(* IEC 61131-3 sources: teller/JD_Teller_LC2_V11/Network/Teller, 1 file *)

(* ---- ONE_Teller_Table.st ---- *)
#define OBJECTS_CONFIG

FUNCTION GLOBAL TAB ONE_Teller
-1$UINT, 0$UINT,
0$UINT, 0$UINT,

13$UDINT,
TO_UDINT(3073024365), "Encoder_Inmeten", 0$UINT, 0$UINT, 1$UINT,
TO_UDINT(1689253198), "FileBase", 1$UINT, 0$UINT, 2$UINT,
TO_UDINT(2225119864), "MerkerEx", 1$UINT, 18$UINT, 2$UINT,
TO_UDINT(1903583397), "Ram", 1$UINT, 3$UINT, 16$UINT,
TO_UDINT(933570811), "RAMex", 1$UINT, 16$UINT, 1$UINT,
TO_UDINT(582296389), "SerSend", 1$UINT, 0$UINT, 1$UINT,
TO_UDINT(1018833242), "SIMPULSJE_Teller", 1$UINT, 0$UINT, 1$UINT,
TO_UDINT(1850111279), "String", 1$UINT, 10$UINT, 2$UINT,
TO_UDINT(2898603620), "StringInternal", 1$UINT, 70$UINT, 0$UINT,
TO_UDINT(2685101138), "TanabeCounterSerial", 1$UINT, 0$UINT, 1$UINT,
TO_UDINT(4092741209), "TellerClass_Teller", 1$UINT, 3$UINT, 1$UINT,
TO_UDINT(3232495061), "VirtualBaseInit", 1$UINT, 3$UINT, 0$UINT,
TO_UDINT(589051502), "VisuTeller_Teller", 1$UINT, 0$UINT, 5$UINT,

_NO_ATTR, TO_UDINT(2959661299), "ENCODER_INMETEN1",

_NO_ATTR, TO_UDINT(316419285), "FILEBASE1",
_NO_ATTR, TO_UDINT(2346024303), "FILEBASE2",

1$UINT, TO_UDINT(3025948), "STRING1\MERKEREX0",
1$UINT, TO_UDINT(1480758749), "STRING3\MERKEREX0",

1$UINT, TO_UDINT(4072236793), "SERSEND1\RSELECTOR",
1$UINT, TO_UDINT(3232725082), "TELLERCLASS1\RI2SENCNT",
1$UINT, TO_UDINT(3756668069), "TELLERCLASS1\RIBOXLENGTHCNT",
1$UINT, TO_UDINT(3865050826), "TELLERCLASS1\RIBOXLENGTHJAML",
1$UINT, TO_UDINT(475055017), "TELLERCLASS1\RIBOXLENGTHJAMR",
1$UINT, TO_UDINT(1711364282), "TELLERCLASS1\RIBOXLENGTHJAMSTR",
1$UINT, TO_UDINT(1431716753), "TELLERCLASS1\RIENCDIV",
1$UINT, TO_UDINT(1100143673), "TELLERCLASS1\RIENCMUL",
1$UINT, TO_UDINT(3615109569), "TELLERCLASS1\RISENSORCNT",
1$UINT, TO_UDINT(1331113651), "TELLERCLASS1\RITOTALPRODUCTION",
1$UINT, TO_UDINT(632896864), "TELLERCLASS1\RMINSPOT",
1$UINT, TO_UDINT(1272264235), "TELLERCLASS1\ROCOUNTER",
1$UINT, TO_UDINT(1448788453), "TELLERCLASS1\RSANALOGSPEEDENABLE",
1$UINT, TO_UDINT(3322901645), "TELLERCLASS1\RSEXTRABOX",
1$UINT, TO_UDINT(2626903235), "TELLERCLASS1\RSFACTORANALOGSPEEDIN",
1$UINT, TO_UDINT(2919943508), "TELLERCLASS1\RSMAXSPEED",

_NO_ATTR, TO_UDINT(1200226343), "RAMEX3",

_NO_ATTR, TO_UDINT(2236149643), "SERSEND1",

_NO_ATTR, TO_UDINT(3969721823), "SIMPULSJE5",

_NO_ATTR, TO_UDINT(677614747), "STRING1",
_NO_ATTR, TO_UDINT(3329095095), "STRING3",

_NO_ATTR, TO_UDINT(3886509187), "READ_SERIAL1",

_NO_ATTR, TO_UDINT(326458637), "TELLERCLASS1",

_NO_ATTR, TO_UDINT(2767617665), "VISUTELLER1",
_NO_ATTR, TO_UDINT(1040133947), "VISUTELLER2",
_NO_ATTR, TO_UDINT(1257775021), "VISUTELLER3",
_NO_ATTR, TO_UDINT(3567028750), "VISUTELLER4",
_NO_ATTR, TO_UDINT(2744892056), "VISUTELLER5",

//Internal connections
0$UDINT,
18$UDINT,
TO_UDINT(22), "rSelector", TO_UDINT(5),
TO_UDINT(24), "MerkerEx0", TO_UDINT(3),
TO_UDINT(25), "MerkerEx0", TO_UDINT(4),
TO_UDINT(27), "RMinSpot", TO_UDINT(15),
TO_UDINT(27), "rSextraBox", TO_UDINT(18),
TO_UDINT(27), "riEncMul", TO_UDINT(12),
TO_UDINT(27), "riEncDiv", TO_UDINT(11),
TO_UDINT(27), "riSensorCNT", TO_UDINT(13),
TO_UDINT(27), "riBoxlengthCNT", TO_UDINT(7),
TO_UDINT(27), "riTotalProduction", TO_UDINT(14),
TO_UDINT(27), "riBoxlengthJAML", TO_UDINT(8),
TO_UDINT(27), "riBoxlengthJAMR", TO_UDINT(9),
TO_UDINT(27), "riBoxlengthJamSTR", TO_UDINT(10),
TO_UDINT(27), "roCounter", TO_UDINT(16),
TO_UDINT(27), "ri2SenCNT", TO_UDINT(6),
TO_UDINT(27), "rsMaxSpeed", TO_UDINT(20),
TO_UDINT(27), "rsFactorAnalogSpeedIn", TO_UDINT(19),
TO_UDINT(27), "rsAnalogSpeedEnable", TO_UDINT(17),
0$UDINT,
27$UDINT,
TO_UDINT(22), "fb", TO_UDINT(1), "Server0",
TO_UDINT(22), "strSend", TO_UDINT(25), "Data",
TO_UDINT(24), "DataBuffer", TO_UDINT(3), "m_udLength",
TO_UDINT(25), "DataBuffer", TO_UDINT(4), "m_udLength",
TO_UDINT(26), "GetInfo", TO_UDINT(27), "ClassSvr",
TO_UDINT(26), "String", TO_UDINT(24), "Data",
TO_UDINT(26), "FileBase", TO_UDINT(2), "Server0",
TO_UDINT(26), "cPlannedProduction", TO_UDINT(27), "iTotalProduction",
TO_UDINT(26), "cBoxLength", TO_UDINT(27), "iBoxlengthCNT",
TO_UDINT(26), "cBattingStart", TO_UDINT(30), "iStart",
TO_UDINT(26), "cBattingDistance", TO_UDINT(30), "iLengte",
TO_UDINT(26), "cBatch1", TO_UDINT(30), "iPakket1SET",
TO_UDINT(26), "cBatch2", TO_UDINT(30), "iPakket2SET",
TO_UDINT(26), "cStartingDistanceToConveyorRun", TO_UDINT(29), "iLengte",
TO_UDINT(26), "cCountedBoxes", TO_UDINT(27), "oCounter",
TO_UDINT(27), "RamEx", TO_UDINT(21), "m_udLength",
TO_UDINT(27), "iSimPuls", TO_UDINT(23), "Uitgang",
TO_UDINT(27), "coTotalproduction", TO_UDINT(22), "iTotalproduction",
TO_UDINT(27), "coCounter", TO_UDINT(22), "iCounter",
TO_UDINT(27), "coRemainingproduction", TO_UDINT(22), "iRemaningproduction",
TO_UDINT(27), "coCounterPerMin", TO_UDINT(22), "iCounterPerMin",
TO_UDINT(27), "coSpeed", TO_UDINT(22), "iSpeed",
TO_UDINT(28), "cData", TO_UDINT(27), "sData",
TO_UDINT(29), "cData", TO_UDINT(27), "sData",
TO_UDINT(30), "cData", TO_UDINT(27), "sData",
TO_UDINT(31), "cData", TO_UDINT(27), "sData",
TO_UDINT(32), "cData", TO_UDINT(27), "sData",

//Initialization values
0$UDINT,
19$UDINT,
TO_UDINT(0), "cEncoder", TO_UDINT(0),//|Teller.Encoder_Inmeten1.cEncoder;
TO_UDINT(3), "ThreadSafe", TO_UDINT(0),//|Teller.String1\MerkerEx0.ThreadSafe;
TO_UDINT(4), "ThreadSafe", TO_UDINT(0),//|Teller.String3\MerkerEx0.ThreadSafe;
TO_UDINT(21), "ThreadSafe", TO_UDINT(0),//|Teller.RAMex3.ThreadSafe;
TO_UDINT(24), "SingleRealloc", TO_UDINT(1),//|Teller.String1.SingleRealloc;
TO_UDINT(26), "GetInfo", TO_UDINT(0),//|Teller.Read_serial1.GetInfo;
TO_UDINT(27), "iSensorSTR", TO_UDINT(0),//|Teller.TellerClass1.iSensorSTR;
TO_UDINT(27), "oJam", TO_UDINT(0),//|Teller.TellerClass1.oJam;
TO_UDINT(27), "cExtBoxCount", TO_UDINT(0),//|Teller.TellerClass1.cExtBoxCount;
TO_UDINT(28), "cHeadNr", TO_UDINT(1),//|Teller.VisuTeller1.cHeadNr;
TO_UDINT(28), "cType", TO_UDINT(4),//|Teller.VisuTeller1.cType;
TO_UDINT(29), "cHeadNr", TO_UDINT(2),//|Teller.VisuTeller2.cHeadNr;
TO_UDINT(29), "cType", TO_UDINT(3),//|Teller.VisuTeller2.cType;
TO_UDINT(30), "cHeadNr", TO_UDINT(3),//|Teller.VisuTeller3.cHeadNr;
TO_UDINT(30), "cType", TO_UDINT(1),//|Teller.VisuTeller3.cType;
TO_UDINT(31), "cHeadNr", TO_UDINT(4),//|Teller.VisuTeller4.cHeadNr;
TO_UDINT(31), "cType", TO_UDINT(5),//|Teller.VisuTeller4.cType;
TO_UDINT(32), "cHeadNr", TO_UDINT(5),//|Teller.VisuTeller5.cHeadNr;
TO_UDINT(32), "cType", TO_UDINT(2),//|Teller.VisuTeller5.cType;

//Symbolic initialization values
0$UDINT,
0$UDINT,

//Initialization of string values
0$UDINT,
0$UDINT,

//Configuration of tasks (RealTime, Cyclic, Background)
0$UDINT,
1$UDINT,
TO_UDINT(27), (1)$UDINT, 4194305$DINT, 	//TELLERCLASS1

0$UDINT,
3$UDINT,
TO_UDINT(26), (1)$UDINT, 4194303$DINT, 	//READ_SERIAL1
TO_UDINT(23), (10)$UDINT, 4194305$DINT, 	//SIMPULSJE5
TO_UDINT(27), (100)$UDINT, 4194305$DINT, 	//TELLERCLASS1

0$UDINT,
6$UDINT,
TO_UDINT(27), (200)$UDINT, 4194305$DINT, 	//TELLERCLASS1
TO_UDINT(28), (200)$UDINT, 4194305$DINT, 	//VISUTELLER1
TO_UDINT(29), (200)$UDINT, 4194305$DINT, 	//VISUTELLER2
TO_UDINT(30), (200)$UDINT, 4194305$DINT, 	//VISUTELLER3
TO_UDINT(31), (200)$UDINT, 4194305$DINT, 	//VISUTELLER4
TO_UDINT(32), (200)$UDINT, 4194305$DINT, 	//VISUTELLER5

//External connections
0$UDINT,
15$UDINT,
TO_UDINT(0), "cEncoder", C_DIR, TO_UDINT(396609901), "CIO011_IM1","Encoder",
TO_UDINT(22), "Ser", C_DIR, TO_UDINT(2650501396), "CIV5211\_VaranSerLibOS0","Command",
TO_UDINT(26), "RxTx", C_DIR, TO_UDINT(3942400386), "CIV5211\_VaranSerLibOS1","Command",
TO_UDINT(27), "iEncoder", C_TRY, TO_UDINT(396609901), "CIO011_IM1","Encoder",
TO_UDINT(27), "iSensorL", C_TRY, TO_UDINT(396609901), "CIO011_IM1","Input4",
TO_UDINT(27), "iSensorR", C_TRY, TO_UDINT(396609901), "CIO011_IM1","Input5",
TO_UDINT(27), "iSensorSTR", C_TRY, TO_UDINT(396609901), "CIO011_IM1","Input3",
TO_UDINT(27), "oHeadnr01", C_TRY, TO_UDINT(396609901), "CIO011_IM1","Output4",
TO_UDINT(27), "oHeadnr02", C_TRY, TO_UDINT(396609901), "CIO011_IM1","Output5",
TO_UDINT(27), "oHeadnr03", C_TRY, TO_UDINT(396609901), "CIO011_IM1","Output2",
TO_UDINT(27), "oHeadnr04", C_TRY, TO_UDINT(396609901), "CIO011_IM1","Output1",
TO_UDINT(27), "oHeadnr05", C_TRY, TO_UDINT(396609901), "CIO011_IM1","Output3",
TO_UDINT(27), "c_JamData", C_DIR, TO_UDINT(2288677303), "S11_RAM_Jamdetection_TeachIn_01","m_udLength",
TO_UDINT(27), "cAnalogSpeedOut", C_DIR, TO_UDINT(396609901), "CIO011_IM1","AO",
TO_UDINT(27), "cExtBoxCount", C_DIR, TO_UDINT(396609901), "CIO011_IM1","Output7",

//Magic internal connections
0$UDINT,
0$UDINT,

//Configuration of timeslots of tasks (RealTime, Cyclic)
#ifdef __LSLLDR_TIMESLOTS__
0$UDINT,
0$UDINT,

0$UDINT,
0$UDINT,

#endif //__LSLLDR_TIMESLOTS__

//MultiMaster connections
#ifdef __LSLLDR_MULTIMASTER__
0$UDINT,
0$UDINT,
#endif //__LSLLDR_MULTIMASTER__

END_FUNCTION
